Fanuc KAREL source: ka00144.KL

-- PROVISIONAL review KL for V770-1; original PC SHA256 d511f9396c269090f3b8e1e23180439a83cff972449fac5734c05dfc7be255b6
-- Incomplete behavior may be omitted. Consult companion uncertainty JSON. Do not deploy.
PROGRAM KA00144
%NOLOCKGROUP
-- UNRESOLVED_DECL SRC type=002017
-- UNRESOLVED_DECL DST type=002017
BEGIN
  -- UNRESOLVED_PC offsets 5-19; opcodes 2E,22,9D,33,B4
  -- UNRESOLVED_PC offsets 24-42; opcodes 22,9D,33,B3,22,9D,33,B4
  -- UNRESOLVED_PC offsets 47-51; opcodes 7F
END KA00144
